// TIA Portal V15.1 export
DATA_BLOCK "MCP_RC_R5DBB"   // DB9831
{ S7_Optimized_Access := 'TRUE' }
   VAR
      Motor : "MCP_RC_R5UDT";
      Level : Int := 7;
   END_VAR
BEGIN
   Motor.Speed := 2.5;
END_DATA_BLOCK
